FUNCTION_BLOCK MOD_StateLogic (* The PackML state machine itself: Reset, Start, Stop, Abort and Clear take it from state to state (MOD_StateGate has already checked who sent them, and that PackML allows them now); while Stopping it waits until no skill runs any more. Technical: PackML module state machine: RESET, START, STOP, ABORT, CLEAR (decided by MOD_StateGate); runs the Resetting and Stopping procedures; Stopping waits until no skill is active *)
  (* Standard: 61499-2 *)
  (* Version 0.1, 2026-09-28, Project contributors, AAU Smart Production Lab *)
  PACKAGE modlib;
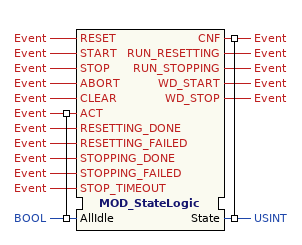
  EVENT_INPUT
    RESET; (* Reset the module (accepted by MOD_StateGate) *)
    START; (* Start the module (accepted by MOD_StateGate) *)
    STOP; (* Stop the module (accepted by MOD_StateGate) *)
    ABORT; (* Abort the module (accepted by MOD_StateGate) *)
    CLEAR; (* Clear the module (accepted by MOD_StateGate) *)
    ACT WITH AllIdle; (* The number of running skills changed (AllIdle) *)
    RESETTING_DONE; (* The Resetting procedure ended *)
    RESETTING_FAILED; (* The Resetting procedure failed *)
    STOPPING_DONE; (* The Stopping procedure ended *)
    STOPPING_FAILED; (* The Stopping procedure failed *)
    STOP_TIMEOUT; (* Stopping took longer than StopTimeout *)
  END_EVENT
  EVENT_OUTPUT
    CNF WITH State; (* The state changed *)
    RUN_RESETTING; (* Run the Resetting procedure *)
    RUN_STOPPING; (* Run the Stopping procedure *)
    WD_START; (* Start the stop timeout *)
    WD_STOP; (* Stop the stop timeout *)
  END_EVENT
  VAR_INPUT
    AllIdle : BOOL := TRUE; (* No skill runs *)
  END_VAR
  VAR_OUTPUT
    State : USINT := 2; (* PackML state: 1 Clearing, 2 Stopped, 3 Starting, 4 Idle, 6 Execute, 7 Stopping, 8 Aborting, 9 Aborted, 15 Resetting *)
  END_VAR
  EC_STATES
    Stopped : Alg_Stopped -> CNF;
    Resetting : Alg_Resetting -> CNF, -> RUN_RESETTING;
    ResettingW;
    Idle : Alg_Idle -> CNF;
    Starting : Alg_Starting -> CNF;
    Execute : Alg_Execute -> CNF;
    Stopping : Alg_Stopping -> CNF, -> WD_START;
    StoppingW;
    StopProc : -> WD_STOP, -> RUN_STOPPING;
    StopProcW;
    Aborting : Alg_Aborting -> CNF, -> WD_STOP;
    Aborted : Alg_Aborted -> CNF;
    Clearing : Alg_Clearing -> CNF;
  END_STATES
  EC_TRANSITIONS
    Stopped TO Resetting := RESET;
    Idle TO Starting := START;
    ResettingW TO Stopping := STOP;
    Idle TO Stopping := STOP;
    Execute TO Stopping := STOP;
    Stopped TO Aborting := ABORT;
    ResettingW TO Aborting := ABORT;
    Idle TO Aborting := ABORT;
    Execute TO Aborting := ABORT;
    StoppingW TO Aborting := ABORT;
    StopProcW TO Aborting := ABORT;
    Aborted TO Clearing := CLEAR;
    Resetting TO ResettingW := 1;
    ResettingW TO Idle := RESETTING_DONE;
    ResettingW TO Aborting := RESETTING_FAILED;
    Starting TO Execute := 1;
    Stopping TO StoppingW := 1;
    StoppingW TO StopProc := [AllIdle];
    StoppingW TO Aborting := STOP_TIMEOUT;
    StopProc TO StopProcW := 1;
    StopProcW TO Stopped := STOPPING_DONE;
    StopProcW TO Aborting := STOPPING_FAILED;
    Aborting TO Aborted := 1;
    Clearing TO Stopped := 1;
  END_TRANSITIONS
  ALGORITHM Alg_Stopped IN ST:
State := 2;
  END_ALGORITHM
  ALGORITHM Alg_Resetting IN ST:
State := 15;
  END_ALGORITHM
  ALGORITHM Alg_Idle IN ST:
State := 4;
  END_ALGORITHM
  ALGORITHM Alg_Starting IN ST:
State := 3;
  END_ALGORITHM
  ALGORITHM Alg_Execute IN ST:
State := 6;
  END_ALGORITHM
  ALGORITHM Alg_Stopping IN ST:
State := 7;
  END_ALGORITHM
  ALGORITHM Alg_Aborting IN ST:
State := 8;
  END_ALGORITHM
  ALGORITHM Alg_Aborted IN ST:
State := 9;
  END_ALGORITHM
  ALGORITHM Alg_Clearing IN ST:
State := 1;
  END_ALGORITHM
END_FUNCTION_BLOCK
